// TIA Portal V20 export
// export: Created 2026-10-12T16:46:22.7383713Z, ExportSetting WithDefaults, DisplayName Totally Integrated Automation Portal, DisplayVersion V20 Update 6, DisplayName TIA Portal Openness, DisplayVersion V20 Update 6, DisplayName TIA Portal Version Control Interface, DisplayVersion V20 Update 6, DisplayName SINAMICS Startdrive Advanced, DisplayVersion V20 SP1 Update 2, DisplayName SINAMICS Startdrive G110M, G120, G120C, G120D, G120P, G115D, DisplayVersion V20 SP1 Update 2, DisplayName SINAMICS Startdrive G130, G150, S120, S150, SINAMICS MV, G220, S200, S210, DisplayVersion V20 SP1 Update 2, DisplayName STEP 7 Professional, DisplayVersion V20 Update 6, DisplayName STEP 7 Safety, DisplayVersion V20 Update 2, DisplayName WinCC Basic/Comfort/Advanced, DisplayVersion V20 Update 6, DisplayName WinCC Professional, DisplayVersion V20 Update 6, DisplayName WinCC Unified, DisplayVersion V20 Update 6
TYPE "UDT_FlexKraft_In"
// ==============================================================================
//  UDT 2: Input  (FK Input Register 0..15 -> Gateway -> SPS)
// ==============================================================================
// stored: IsFailsafeCompliant false
   STRUCT
      Reserved0 : Word;   // Reg 0 immer 16#0000
      StatusRegister : Word;   // Reg 1 Bitfeld
      WarningsRegister : Word;   // Reg 2 Bitfeld
      AlarmsRegister : Word;   // Reg 3 Bitfeld
      OutputVoltage : Int;   // Reg 4 Istspannung *0,01 V
      OutputCurrent : Int;   // Reg 5 Iststrom *1 A bzw. *0,1 A (HiRes)
      ProcessTime_HW : Word;   // Reg 6
      ProcessTime_LW : Word;   // Reg 7
      Ah_HW : Word;   // Reg 8
      Ah_LW : Word;   // Reg 9
      Reserved : Array[10..15] of Word;   // Reg 10..15 ungenutzt
   END_STRUCT;
END_TYPE
